fbExtDisableAF(
    Axis := axis3,
    Execute := bForceFall OR bEStopActive OR bNeedAxisReset
);

fbExtDisableYaw(
    Axis := axis4,
    Execute := bForceFall OR bEStopActive OR bNeedAxisReset
);

bExtBD := fbExtEnableBD.Enabled;
bExtAC := fbExtEnableAC.Enabled;
bExtAF := fbExtEnableAF.Enabled;
bExtYaw := fbExtEnableYaw.Enabled;

bRunForce := bForceMode
             AND bZeroDone
             AND bAxesReadyForForce
             AND axis1_power.Status
             AND Axis1_BrakeMotionOK
             AND axis2_power.Status
             AND axis3_power.Status
             AND axis4_power.Status
             AND bExtBD
             AND bExtAC
             AND bExtAF
             AND bExtYaw;

// 未进入实际力控运行（包括退出、急停、轴未就绪）时清除平面历史意图。
IF NOT bRunForce THEN
    bXIntent := FALSE;
    bZIntent := FALSE;
    bXDriveActive := FALSE;
    bZDriveActive := FALSE;
    Fx_work_target := 0.0;
    Fz_work_target := 0.0;
    Fx_work := 0.0;
    Fz_work := 0.0;
END_IF;


// =============================================================
// O. 编码器值 -> 机构学位置
// AC：-59 编码器对应 90°，编码器增大角度减小
// =============================================================
LBD_mm := BD_ActEnc + BD_KinOffset_mm;
LBD_m  := LBD_mm / 1000.0;

ThetaAC_deg := AC_ThetaRef_deg - (AC_ActEnc - AC_EncRef_deg);
ThetaAC_rad := ThetaAC_deg * DEG2RAD;


// =============================================================
// P. 当前 E 点正解
// =============================================================
bGeoOK := FALSE;

Cx := Ax0 + l_AC * COS(ThetaAC_rad);
Cz := Az0 + l_AC * SIN(ThetaAC_rad);

dxBC := Cx - Bx0;
dzBC := Cz - Bz0;
dBC := SQRT(dxBC * dxBC + dzBC * dzBC);

IF (LBD_m > 0.01) AND (dBC > 0.01) THEN
    IF (dBC < (LBD_m + l_CD - GeoMargin_m)) AND
       (dBC > (ABS(LBD_m - l_CD) + GeoMargin_m)) THEN

        alphaBC := F_Atan2_LREAL(y := dzBC, x := dxBC);
        cosBeta := (LBD_m * LBD_m + dBC * dBC - l_CD * l_CD) / (2.0 * LBD_m * dBC);

        IF (cosBeta <= 1.0) AND (cosBeta >= -1.0) THEN
            beta := ACOS(cosBeta);
            thBD := alphaBC - beta;

            Dx := Bx0 + LBD_m * COS(thBD);
            Dz := Bz0 + LBD_m * SIN(thBD);

            theta3 := F_Atan2_LREAL(y := Dz - Cz, x := Dx - Cx);

            // D 点不在 CE 上：D 相对 CE 垂直偏置 D_Offset_m
            // theta3 是 CD 方向，thetaCE 才是 CE 主杆方向
            IF l_CD > D_Offset_m THEN
                s_CD_CE := SQRT(l_CD * l_CD - D_Offset_m * D_Offset_m);
                gamma_DCE := ATAN(D_Offset_m / s_CD_CE);
                thetaCE := theta3 + CE_Sign * gamma_DCE;

                Ex := Cx + l_CE * COS(thetaCE);
                Ez := Cz + l_CE * SIN(thetaCE);

                bGeoOK := TRUE;
            END_IF;
        END_IF;
    END_IF;
END_IF;


// =============================================================
// Q. AC 机构角扰动 E 点正解
// =============================================================
bGeoOK_th := FALSE;

Cx_th := Ax0 + l_AC * COS(ThetaAC_rad + dTheta);
Cz_th := Az0 + l_AC * SIN(ThetaAC_rad + dTheta);

dxBC_th := Cx_th - Bx0;
dzBC_th := Cz_th - Bz0;
dBC_th := SQRT(dxBC_th * dxBC_th + dzBC_th * dzBC_th);

IF (LBD_m > 0.01) AND (dBC_th > 0.01) THEN
    IF (dBC_th < (LBD_m + l_CD - GeoMargin_m)) AND
       (dBC_th > (ABS(LBD_m - l_CD) + GeoMargin_m)) THEN

        alphaBC_th := F_Atan2_LREAL(y := dzBC_th, x := dxBC_th);
        cosBeta_th := (LBD_m * LBD_m + dBC_th * dBC_th - l_CD * l_CD) / (2.0 * LBD_m * dBC_th);

        IF (cosBeta_th <= 1.0) AND (cosBeta_th >= -1.0) THEN
            beta_th := ACOS(cosBeta_th);
            thBD_th := alphaBC_th - beta_th;

            Dx_th := Bx0 + LBD_m * COS(thBD_th);
            Dz_th := Bz0 + LBD_m * SIN(thBD_th);

            theta3_th := F_Atan2_LREAL(y := Dz_th - Cz_th, x := Dx_th - Cx_th);

            IF l_CD > D_Offset_m THEN
                s_CD_CE_th := SQRT(l_CD * l_CD - D_Offset_m * D_Offset_m);
                gamma_DCE_th := ATAN(D_Offset_m / s_CD_CE_th);
                thetaCE_th := theta3_th + CE_Sign * gamma_DCE_th;

                Ex_th := Cx_th + l_CE * COS(thetaCE_th);
                Ez_th := Cz_th + l_CE * SIN(thetaCE_th);

                bGeoOK_th := TRUE;
            END_IF;
        END_IF;
    END_IF;
END_IF;


// =============================================================
// R. BD 机构长度扰动 E 点正解
// =============================================================
bGeoOK_L := FALSE;

Cx_L := Cx;
Cz_L := Cz;

dxBC_L := Cx_L - Bx0;
dzBC_L := Cz_L - Bz0;
dBC_L := SQRT(dxBC_L * dxBC_L + dzBC_L * dzBC_L);

IF ((LBD_m + dL) > 0.01) AND (dBC_L > 0.01) THEN
    IF (dBC_L < ((LBD_m + dL) + l_CD - GeoMargin_m)) AND
       (dBC_L > (ABS((LBD_m + dL) - l_CD) + GeoMargin_m)) THEN

        alphaBC_L := F_Atan2_LREAL(y := dzBC_L, x := dxBC_L);
        cosBeta_L := ((LBD_m + dL) * (LBD_m + dL) + dBC_L * dBC_L - l_CD * l_CD)
                     / (2.0 * (LBD_m + dL) * dBC_L);

        IF (cosBeta_L <= 1.0) AND (cosBeta_L >= -1.0) THEN
            beta_L := ACOS(cosBeta_L);
            thBD_L := alphaBC_L - beta_L;

            Dx_L := Bx0 + (LBD_m + dL) * COS(thBD_L);
            Dz_L := Bz0 + (LBD_m + dL) * SIN(thBD_L);

            theta3_L := F_Atan2_LREAL(y := Dz_L - Cz_L, x := Dx_L - Cx_L);

            IF l_CD > D_Offset_m THEN
                s_CD_CE_L := SQRT(l_CD * l_CD - D_Offset_m * D_Offset_m);
                gamma_DCE_L := ATAN(D_Offset_m / s_CD_CE_L);
                thetaCE_L := theta3_L + CE_Sign * gamma_DCE_L;

                Ex_L := Cx_L + l_CE * COS(thetaCE_L);
                Ez_L := Cz_L + l_CE * SIN(thetaCE_L);

                bGeoOK_L := TRUE;
            END_IF;
        END_IF;
    END_IF;
END_IF;


// =============================================================
// S. E 点速度雅可比
// =============================================================
bValidJ := FALSE;
bSingular := FALSE;

IF bGeoOK AND bGeoOK_th AND bGeoOK_L THEN
    J11 := (Ex_th - Ex) / dTheta;
    J21 := (Ez_th - Ez) / dTheta;

    J12 := (Ex_L - Ex) / dL;
    J22 := (Ez_L - Ez) / dL;

    detJ := J11 * J22 - J12 * J21;

    IF ABS(detJ) > DetMin THEN
        bValidJ := TRUE;
    ELSE
        bSingular := TRUE;
    END_IF;
END_IF;


// =============================================================
// T. AC/BD 二维导纳 + 雅可比逆解
// 1) 平面 X/Z 导纳由显式欧拉改为一阶精确离散：M * dV/dt + B * V = F
//    Vss = Fadm / B
//    V(k+1) = Vss + (V(k)-Vss) * EXP(-B*Ts/M)
// 2) 撤力时使用 AdmB_Stop_X/Z 平滑衰减，轴减速度限幅约束最终命令。
// 3) VxyMax_mps = 0.300，先限制末端合速度，再做 J^-1。
// =============================================================
BD_Vraw_enc_s := 0.0;
AC_Vraw_enc_s := 0.0;
AF_Vraw_enc_s := 0.0;
Yaw_Vraw_enc_s := 0.0;

IF bRunForce AND bValidJ THEN
    Vx_last_mps := Vx_mps;
    Vz_last_mps := Vz_mps;

    // X 通道：有力用运动阻尼，撤力用停车阻尼。
    IF NOT bXDriveActive THEN
        AdmB_Use_X := AdmB_Stop_X;
        Fadm_X := 0.0;
    ELSE
        AdmB_Use_X := AdmB_Move_X;
        Fadm_X := ForceGain_X * TransWeight_X * Fx_work;
    END_IF;

    // Z 通道：有力用运动阻尼，撤力用停车阻尼。
    IF NOT bZDriveActive THEN
        AdmB_Use_Z := AdmB_Stop_Z;
        Fadm_Z := 0.0;
    ELSE
        AdmB_Use_Z := AdmB_Move_Z;
        Fadm_Z := ForceGain_Z * TransWeight_Z * Fz_work;
    END_IF;

    // M/B 安全保护，防止除零或负值。
    IF AdmM_X < 0.001 THEN
        AdmM_X_Use := 0.001;
    ELSE
        AdmM_X_Use := AdmM_X;
    END_IF;

    IF AdmM_Z < 0.001 THEN
        AdmM_Z_Use := 0.001;
    ELSE
        AdmM_Z_Use := AdmM_Z;
    END_IF;

    IF AdmB_Use_X < 0.001 THEN
        AdmB_X_UseSafe := 0.001;
    ELSE
        AdmB_X_UseSafe := AdmB_Use_X;
    END_IF;

    IF AdmB_Use_Z < 0.001 THEN
        AdmB_Z_UseSafe := 0.001;
    ELSE
        AdmB_Z_UseSafe := AdmB_Use_Z;
    END_IF;

    // 稳态速度。撤力时 Fadm=0，因此 Vss=0。
    Vxss_mps := Fadm_X / AdmB_X_UseSafe;
    Vzss_mps := Fadm_Z / AdmB_Z_UseSafe;

    // 精确离散指数项。
    IF Ts > 0.000001 THEN
        Vx_ExpK := EXP(-AdmB_X_UseSafe * Ts / AdmM_X_Use);
        Vz_ExpK := EXP(-AdmB_Z_UseSafe * Ts / AdmM_Z_Use);
    ELSE
        Vx_ExpK := 0.0;
        Vz_ExpK := 0.0;
    END_IF;

    Vx_mps := Vxss_mps + (Vx_last_mps - Vxss_mps) * Vx_ExpK;
    Vz_mps := Vzss_mps + (Vz_last_mps - Vzss_mps) * Vz_ExpK;

    IF Ts > 0.000001 THEN
        Ax_mps2 := (Vx_mps - Vx_last_mps) / Ts;
        Az_mps2 := (Vz_mps - Vz_last_mps) / Ts;
    ELSE
        Ax_mps2 := 0.0;
        Az_mps2 := 0.0;
    END_IF;

    // NaN / 极大值保护，避免后续 J^-1 或限幅触发 FPU invalid。
    IF Vx_mps <> Vx_mps THEN
        Vx_mps := 0.0;
        Vx_last_mps := 0.0;
        Ax_mps2 := 0.0;
    ELSIF ABS(Vx_mps) > Vplane_NumLimit_mps THEN
        Vx_mps := 0.0;
        Vx_last_mps := 0.0;
        Ax_mps2 := 0.0;
    END_IF;

    IF Vz_mps <> Vz_mps THEN
        Vz_mps := 0.0;
        Vz_last_mps := 0.0;
        Az_mps2 := 0.0;
    ELSIF ABS(Vz_mps) > Vplane_NumLimit_mps THEN
        Vz_mps := 0.0;
        Vz_last_mps := 0.0;
        Az_mps2 := 0.0;
    END_IF;

    // 限幅前理论平面速度。
    Vnorm_PreLimit_mps := SQRT(Vx_mps * Vx_mps + Vz_mps * Vz_mps);

    IF Vnorm_PreLimit_mps > VxyMax_mps THEN
        ScaleVel_Plane := VxyMax_mps / Vnorm_PreLimit_mps;
        Vx_mps := Vx_mps * ScaleVel_Plane;
        Vz_mps := Vz_mps * ScaleVel_Plane;
    ELSE
        ScaleVel_Plane := 1.0;
    END_IF;

    // 限幅后的真实平面速度。Watch 中 Vnorm 显示这个值。
    Vnorm_AfterLimit_mps := SQRT(Vx_mps * Vx_mps + Vz_mps * Vz_mps);
    Vnorm := Vnorm_AfterLimit_mps;

    qdotAC_rad_s := ( J22 * Vx_mps - J12 * Vz_mps) / detJ;
    qdotBD_m_s   := (-J21 * Vx_mps + J11 * Vz_mps) / detJ;

    // AC：机构角增大时，编码器减小。
    AC_Vraw_enc_s := -qdotAC_rad_s * RAD2DEG;

    // BD：1 mm = 1 mm，不做比例换算。
    BD_Vraw_enc_s := qdotBD_m_s * 1000.0;

ELSE
    Vx_mps := 0.0;
    Vz_mps := 0.0;
    Vx_last_mps := 0.0;
    Vz_last_mps := 0.0;

    Ax_mps2 := 0.0;
    Az_mps2 := 0.0;

    Vnorm_PreLimit_mps := 0.0;
    Vnorm_AfterLimit_mps := 0.0;
    Vnorm := 0.0;
    ScaleVel_Plane := 1.0;

    qdotAC_rad_s := 0.0;
    qdotBD_m_s := 0.0;
END_IF;

// axis3 AF 俯仰：Tz/Mz -> 俯仰角速度
// 本版关键修改：
// 1) 不再用显式欧拉 W += ((Madm-B*W)/J)*Ts 处理大 Stop 阻尼；
// 2) 改用一阶系统精确离散 W_new = Wss + (W_old-Wss)*EXP(-B*Ts/J)；
// 3) 撤力阻尼保持温和，减速由 AF_Dmax_enc_s2 最终约束。
IF bRunForce THEN
    AF_W_last_enc_s := AF_W_enc_s;

    bAF_TorqueActive := ABS(Mz_work_Nm) > 0.0001;

    IF bAF_TorqueActive THEN
        AdmB_Use_AF := AdmB_Move_AF;
        Madm_AF := TorqueGain_AF * Dir_Mz_AF * Mz_work_Nm;
    ELSE
        AdmB_Use_AF := AdmB_Stop_AF;
        Madm_AF := 0.0;
    END_IF;

    // 数值保护：J 和 B 都不允许过小。
    IF AdmJ_AF < 0.001 THEN
        AdmJ_AF_Use := 0.001;
    ELSE
        AdmJ_AF_Use := AdmJ_AF;
    END_IF;

    IF AdmB_Use_AF < 0.001 THEN
        AdmB_AF_UseSafe := 0.001;
    ELSE
        AdmB_AF_UseSafe := AdmB_Use_AF;
    END_IF;

    // 一阶导纳精确离散，撤力阻尼决定内部角速度衰减时间常数。
    IF Ts > 0.000001 THEN
        AF_ExpK := EXP(-AdmB_AF_UseSafe * Ts / AdmJ_AF_Use);
    ELSE
        AF_ExpK := 0.0;
    END_IF;

    AF_Wss_enc_s := Madm_AF / AdmB_AF_UseSafe;
    AF_W_enc_s := AF_Wss_enc_s + (AF_W_last_enc_s - AF_Wss_enc_s) * AF_ExpK;

    // 撤力后小速度直接归零，避免低速漂移。
    IF (NOT bAF_TorqueActive) AND (ABS(AF_W_enc_s) < AF_StopZeroVel_enc_s) THEN
        AF_W_enc_s := 0.0;
    END_IF;

    IF Ts > 0.000001 THEN
        AF_Alpha_enc_s2 := (AF_W_enc_s - AF_W_last_enc_s) / Ts;
    ELSE
        AF_Alpha_enc_s2 := 0.0;
    END_IF;

    // NaN / 极大值保护，避免再次触发 FPU invalid。
    IF AF_W_enc_s <> AF_W_enc_s THEN
        AF_W_enc_s := 0.0;
        AF_W_last_enc_s := 0.0;
        AF_Alpha_enc_s2 := 0.0;
    ELSIF ABS(AF_W_enc_s) > AF_NumLimit_enc_s THEN
        AF_W_enc_s := 0.0;
        AF_W_last_enc_s := 0.0;
        AF_Alpha_enc_s2 := 0.0;
    END_IF;

    AF_Vraw_enc_s := AF_W_enc_s;
ELSE
    AF_W_enc_s := 0.0;
    AF_W_last_enc_s := 0.0;
    AF_Alpha_enc_s2 := 0.0;
    AF_Vraw_enc_s := 0.0;
END_IF;

// axis4 底盘 yaw：稳定离散导纳
// 当前 yaw 主输入来自 FzYaw_work_N -> Myaw_work_Nm -> Mx_work_Nm。
// 这里继续使用 Mx_work_Nm 作为 yaw 有效输入，兼容你前面 Watch 变量。
IF bRunForce THEN
    Yaw_W_last_enc_s := Yaw_W_enc_s;

    YawInput_Nm := Mx_work_Nm;

    // 有 yaw 输入时用运动阻尼；撤力后用停车阻尼。
    IF ABS(YawInput_Nm) <= 0.0001 THEN
        AdmB_Use_Yaw := AdmB_Stop_Yaw;
        Madm_Yaw := 0.0;
    ELSE
        AdmB_Use_Yaw := AdmB_Move_Yaw;
        Madm_Yaw := TorqueGain_Yaw * Dir_Mx_Yaw * YawInput_Nm;
    END_IF;

    // J/B 安全保护。
    IF AdmJ_Yaw < 0.001 THEN
        AdmJ_Yaw_Use := 0.001;
    ELSE
        AdmJ_Yaw_Use := AdmJ_Yaw;
    END_IF;

    IF AdmB_Use_Yaw < 0.001 THEN
        AdmB_Yaw_UseSafe := 0.001;
    ELSE
        AdmB_Yaw_UseSafe := AdmB_Use_Yaw;
    END_IF;

    // 一阶导纳精确离散：
    // dW/dt = (Madm - B*W)/J
    // Wss = Madm/B
    // W(k+1) = Wss + (W(k)-Wss)*EXP(-B*Ts/J)
    Yaw_Wss_enc_s := Madm_Yaw / AdmB_Yaw_UseSafe;

    IF Ts > 0.000001 THEN
        Yaw_ExpK := EXP(-AdmB_Yaw_UseSafe * Ts / AdmJ_Yaw_Use);
    ELSE
        Yaw_ExpK := 0.0;
    END_IF;

    Yaw_W_enc_s :=
        Yaw_Wss_enc_s
      + (Yaw_W_last_enc_s - Yaw_Wss_enc_s) * Yaw_ExpK;

    IF Ts > 0.000001 THEN
        Yaw_Alpha_enc_s2 := (Yaw_W_enc_s - Yaw_W_last_enc_s) / Ts;
    ELSE
        Yaw_Alpha_enc_s2 := 0.0;
    END_IF;

    // NaN / 极大值保护，避免再次触发 FPU invalid。
    IF Yaw_W_enc_s <> Yaw_W_enc_s THEN
        Yaw_W_enc_s := 0.0;
        Yaw_W_last_enc_s := 0.0;
        Yaw_Alpha_enc_s2 := 0.0;
    ELSIF ABS(Yaw_W_enc_s) > Yaw_NumLimit_enc_s THEN
        Yaw_W_enc_s := 0.0;
        Yaw_W_last_enc_s := 0.0;
        Yaw_Alpha_enc_s2 := 0.0;
    END_IF;

    Yaw_Vraw_enc_s := Yaw_W_enc_s;
ELSE
    Yaw_W_enc_s := 0.0;
    Yaw_W_last_enc_s := 0.0;
    Yaw_Alpha_enc_s2 := 0.0;
    Yaw_Vraw_enc_s := 0.0;
END_IF;




// =============================================================
// T1. 机构学限位对力控 Vraw 的拦截
// 放在 U. 轴速度限幅之前；先判断，再进入速度/加速度/位置积分
// =============================================================
bLimitClampPlanar := FALSE;
bLimitClampAF := FALSE;

// BD 只受 CE-HI 限位
IF (BD_Vraw_enc_s > 0.0) AND bCEHI_Block_BD_Pos THEN
    BD_Vraw_enc_s := 0.0;
    bLimitClampPlanar := TRUE;
END_IF;

IF (BD_Vraw_enc_s < 0.0) AND bCEHI_Block_BD_Neg THEN
    BD_Vraw_enc_s := 0.0;
    bLimitClampPlanar := TRUE;
END_IF;

// AC 同时受 CAF 和 CE-HI 限位
IF (AC_Vraw_enc_s > 0.0) AND (bCAF_Block_AC_Pos OR bCEHI_Block_AC_Pos) THEN
    AC_Vraw_enc_s := 0.0;
    bLimitClampPlanar := TRUE;
END_IF;

IF (AC_Vraw_enc_s < 0.0) AND (bCAF_Block_AC_Neg OR bCEHI_Block_AC_Neg) THEN
    AC_Vraw_enc_s := 0.0;
    bLimitClampPlanar := TRUE;
END_IF;

// AF 同时受 CAF 和 CE-HI 限位
IF (AF_Vraw_enc_s > 0.0) AND (bCAF_Block_AF_Pos OR bCEHI_Block_AF_Pos) THEN
    AF_Vraw_enc_s := 0.0;
    bLimitClampAF := TRUE;
END_IF;

IF (AF_Vraw_enc_s < 0.0) AND (bCAF_Block_AF_Neg OR bCEHI_Block_AF_Neg) THEN
    AF_Vraw_enc_s := 0.0;
    bLimitClampAF := TRUE;
END_IF;

// 清导纳内部速度记忆，防止继续顶限位
IF bLimitClampPlanar THEN
    Vx_mps := 0.0;
    Vz_mps := 0.0;
    Vx_last_mps := 0.0;
    Vz_last_mps := 0.0;
    Ax_mps2 := 0.0;
    Az_mps2 := 0.0;
END_IF;

IF bLimitClampAF THEN
    AF_W_enc_s := 0.0;
    AF_W_last_enc_s := 0.0;
    AF_Alpha_enc_s2 := 0.0;
END_IF;


// =============================================================
// U. 轴速度限幅
// =============================================================
ScaleVel := 1.0;
ScaleVel_Axis := 1.0;

IF ABS(BD_Vraw_enc_s) > BD_Vmax_enc_s THEN
    tmpScale := BD_Vmax_enc_s / ABS(BD_Vraw_enc_s);
    IF tmpScale < ScaleVel THEN
        ScaleVel := tmpScale;
    END_IF;
END_IF;

IF ABS(AC_Vraw_enc_s) > AC_Vmax_enc_s THEN
    tmpScale := AC_Vmax_enc_s / ABS(AC_Vraw_enc_s);
    IF tmpScale < ScaleVel THEN
        ScaleVel := tmpScale;
    END_IF;
END_IF;

ScaleVel_Axis := ScaleVel;

BD_Vraw_enc_s := BD_Vraw_enc_s * ScaleVel_Axis;
AC_Vraw_enc_s := AC_Vraw_enc_s * ScaleVel_Axis;

// AF/Yaw 速度限幅：不用 x/ABS(x)，避免 Infinity/Infinity 触发 FPU invalid。
IF AF_Vraw_enc_s <> AF_Vraw_enc_s THEN
    AF_Vraw_enc_s := 0.0;
    AF_W_enc_s := 0.0;
    AF_W_last_enc_s := 0.0;
ELSIF ABS(AF_Vraw_enc_s) > AF_NumLimit_enc_s THEN
    AF_Vraw_enc_s := 0.0;
    AF_W_enc_s := 0.0;
    AF_W_last_enc_s := 0.0;
END_IF;

IF AF_Vraw_enc_s > AF_Vmax_enc_s THEN
    AF_Vraw_enc_s := AF_Vmax_enc_s;
ELSIF AF_Vraw_enc_s < -AF_Vmax_enc_s THEN
    AF_Vraw_enc_s := -AF_Vmax_enc_s;
END_IF;

IF Yaw_Vraw_enc_s <> Yaw_Vraw_enc_s THEN
    Yaw_Vraw_enc_s := 0.0;
    Yaw_W_enc_s := 0.0;
    Yaw_W_last_enc_s := 0.0;
ELSIF ABS(Yaw_Vraw_enc_s) > 100000.0 THEN
    Yaw_Vraw_enc_s := 0.0;
    Yaw_W_enc_s := 0.0;
    Yaw_W_last_enc_s := 0.0;
END_IF;

IF Yaw_Vraw_enc_s > Yaw_Vmax_enc_s THEN
    Yaw_Vraw_enc_s := Yaw_Vmax_enc_s;
ELSIF Yaw_Vraw_enc_s < -Yaw_Vmax_enc_s THEN
    Yaw_Vraw_enc_s := -Yaw_Vmax_enc_s;
END_IF;


// =============================================================
// V. 加速度限幅
// =============================================================
BD_Vlast_enc_s := BD_Vcmd_enc_s;
AC_Vlast_enc_s := AC_Vcmd_enc_s;
AF_Vlast_enc_s := AF_Vcmd_enc_s;
Yaw_Vlast_enc_s := Yaw_Vcmd_enc_s;

// AC/BD 加减速度限幅：
// 1) 加速使用 BD_Amax/AC_Amax；
// 2) 撤力减速或反向使用 BD_Dmax/AC_Dmax；
// 3) 最后用同一个 ScaleAcc_Axis 同步缩放 BD/AC，保持末端方向不被破坏。
BD_dV_enc_s := BD_Vraw_enc_s - BD_Vlast_enc_s;
AC_dV_enc_s := AC_Vraw_enc_s - AC_Vlast_enc_s;

IF (ABS(BD_Vraw_enc_s) < ABS(BD_Vlast_enc_s)) OR (BD_Vraw_enc_s * BD_Vlast_enc_s < 0.0) THEN
    BD_dVmax_enc_s := BD_Dmax_enc_s2 * Ts;
ELSE
    BD_dVmax_enc_s := BD_Amax_enc_s2 * Ts;
END_IF;

IF (ABS(AC_Vraw_enc_s) < ABS(AC_Vlast_enc_s)) OR (AC_Vraw_enc_s * AC_Vlast_enc_s < 0.0) THEN
    AC_dVmax_enc_s := AC_Dmax_enc_s2 * Ts;
ELSE
    AC_dVmax_enc_s := AC_Amax_enc_s2 * Ts;
END_IF;

ScaleAcc := 1.0;
ScaleAcc_Axis := 1.0;

IF ABS(BD_dV_enc_s) > BD_dVmax_enc_s THEN
    IF BD_dVmax_enc_s > 0.0 THEN
        tmpScale := BD_dVmax_enc_s / ABS(BD_dV_enc_s);
    ELSE
        tmpScale := 0.0;
    END_IF;
    IF tmpScale < ScaleAcc THEN
        ScaleAcc := tmpScale;
    END_IF;
END_IF;

IF ABS(AC_dV_enc_s) > AC_dVmax_enc_s THEN
    IF AC_dVmax_enc_s > 0.0 THEN
        tmpScale := AC_dVmax_enc_s / ABS(AC_dV_enc_s);
    ELSE
        tmpScale := 0.0;
    END_IF;
    IF tmpScale < ScaleAcc THEN
        ScaleAcc := tmpScale;
    END_IF;
END_IF;

ScaleAcc_Axis := ScaleAcc;

BD_Vcmd_enc_s := BD_Vlast_enc_s + BD_dV_enc_s * ScaleAcc_Axis;
AC_Vcmd_enc_s := AC_Vlast_enc_s + AC_dV_enc_s * ScaleAcc_Axis;

IF Ts > 0.000001 THEN
    BD_Acmd_enc_s2 := (BD_Vcmd_enc_s - BD_Vlast_enc_s) / Ts;
    AC_Acmd_enc_s2 := (AC_Vcmd_enc_s - AC_Vlast_enc_s) / Ts;
ELSE
    BD_Acmd_enc_s2 := 0.0;
    AC_Acmd_enc_s2 := 0.0;
END_IF;

// AF 加减速度限幅：加速用 AF_Amax，撤力减速/反向用更大的 AF_Dmax。
AF_dV_enc_s := AF_Vraw_enc_s - AF_Vlast_enc_s;

IF (ABS(AF_Vraw_enc_s) < ABS(AF_Vlast_enc_s)) OR (AF_Vraw_enc_s * AF_Vlast_enc_s < 0.0) THEN
    AF_dVmax_enc_s := AF_Dmax_enc_s2 * Ts;
ELSE
    AF_dVmax_enc_s := AF_Amax_enc_s2 * Ts;
END_IF;

IF AF_dV_enc_s > AF_dVmax_enc_s THEN
    AF_dV_enc_s := AF_dVmax_enc_s;
ELSIF AF_dV_enc_s < -AF_dVmax_enc_s THEN
    AF_dV_enc_s := -AF_dVmax_enc_s;
END_IF;

AF_Vcmd_enc_s := AF_Vlast_enc_s + AF_dV_enc_s;

IF Ts > 0.000001 THEN
    AF_Acmd_enc_s2 := (AF_Vcmd_enc_s - AF_Vlast_enc_s) / Ts;
ELSE
    AF_Acmd_enc_s2 := 0.0;
END_IF;

// yaw 加减速度限幅：加速用 Yaw_Amax，撤力减速/反向用 Yaw_Dmax。
Yaw_dV_enc_s := Yaw_Vraw_enc_s - Yaw_Vlast_enc_s;

IF (ABS(Yaw_Vraw_enc_s) < ABS(Yaw_Vlast_enc_s)) OR (Yaw_Vraw_enc_s * Yaw_Vlast_enc_s < 0.0) THEN
    Yaw_dVmax_enc_s := Yaw_Dmax_enc_s2 * Ts;
ELSE
    Yaw_dVmax_enc_s := Yaw_Amax_enc_s2 * Ts;
END_IF;

IF Yaw_dV_enc_s > Yaw_dVmax_enc_s THEN
    Yaw_dV_enc_s := Yaw_dVmax_enc_s;
ELSIF Yaw_dV_enc_s < -Yaw_dVmax_enc_s THEN
    Yaw_dV_enc_s := -Yaw_dVmax_enc_s;
END_IF;

Yaw_Vcmd_enc_s := Yaw_Vlast_enc_s + Yaw_dV_enc_s;

IF Ts > 0.000001 THEN
    Yaw_Acmd_enc_s2 := (Yaw_Vcmd_enc_s - Yaw_Vlast_enc_s) / Ts;
ELSE
    Yaw_Acmd_enc_s2 := 0.0;
END_IF;




// =============================================================
// V1. 机构学限位对力控 Vcmd 的最终保险
// 放在 W. 小速度归零之前，位置积分之前
// =============================================================
// BD
IF (BD_Vcmd_enc_s > 0.0) AND bCEHI_Block_BD_Pos THEN
    BD_Vcmd_enc_s := 0.0;
    BD_Acmd_enc_s2 := 0.0;
END_IF;

IF (BD_Vcmd_enc_s < 0.0) AND bCEHI_Block_BD_Neg THEN
    BD_Vcmd_enc_s := 0.0;
    BD_Acmd_enc_s2 := 0.0;
END_IF;

// AC
IF (AC_Vcmd_enc_s > 0.0) AND (bCAF_Block_AC_Pos OR bCEHI_Block_AC_Pos) THEN
    AC_Vcmd_enc_s := 0.0;
    AC_Acmd_enc_s2 := 0.0;
END_IF;

IF (AC_Vcmd_enc_s < 0.0) AND (bCAF_Block_AC_Neg OR bCEHI_Block_AC_Neg) THEN
    AC_Vcmd_enc_s := 0.0;
    AC_Acmd_enc_s2 := 0.0;
END_IF;

// AF
IF (AF_Vcmd_enc_s > 0.0) AND (bCAF_Block_AF_Pos OR bCEHI_Block_AF_Pos) THEN
    AF_Vcmd_enc_s := 0.0;
    AF_Acmd_enc_s2 := 0.0;
    AF_W_enc_s := 0.0;
    AF_W_last_enc_s := 0.0;
END_IF;

IF (AF_Vcmd_enc_s < 0.0) AND (bCAF_Block_AF_Neg OR bCEHI_Block_AF_Neg) THEN
    AF_Vcmd_enc_s := 0.0;
    AF_Acmd_enc_s2 := 0.0;
    AF_W_enc_s := 0.0;
    AF_W_last_enc_s := 0.0;
END_IF;


// =============================================================
// W. 小速度归零
// =============================================================
IF ABS(BD_Vcmd_enc_s) < 0.001 THEN
    BD_Vcmd_enc_s := 0.0;
END_IF;

IF ABS(AC_Vcmd_enc_s) < 0.001 THEN
    AC_Vcmd_enc_s := 0.0;
END_IF;

IF ABS(AF_Vcmd_enc_s) < 0.02 THEN
    AF_Vcmd_enc_s := 0.0;
END_IF;

IF ABS(Yaw_Vcmd_enc_s) < 0.001 THEN
    Yaw_Vcmd_enc_s := 0.0;
END_IF;

// =============================================================
// W1. 轴1抱闸未释放时冻结 BD 给定
// 防止抱闸合上或释放延时未到时，BD 外部位置继续积分。
// =============================================================
IF NOT Axis1_BrakeMotionOK THEN
    BD_Vraw_enc_s := 0.0;
    BD_Vcmd_enc_s := 0.0;
    BD_Vlast_enc_s := 0.0;
    BD_Acmd_enc_s2 := 0.0;
    qdotBD_m_s := 0.0;
    BD_PosCmd_Enc := BD_ActEnc;
END_IF;


// =============================================================
// X. 力控基础软限位
// 当前只对 axis1=BD 编码器 2~600 做限位
// =============================================================
bForceSoftLimit := FALSE;

BD_NextCmd_Enc := BD_PosCmd_Enc + BD_Vcmd_enc_s * Ts;
AC_NextCmd_Enc := AC_PosCmd_Enc + AC_Vcmd_enc_s * Ts;
AF_NextCmd_Enc := AF_PosCmd_Enc + AF_Vcmd_enc_s * Ts;
Yaw_NextCmd_Enc := Yaw_PosCmd_Enc + Yaw_Vcmd_enc_s * Ts;

IF (BD_NextCmd_Enc < BD_EncMin) OR (BD_NextCmd_Enc > BD_EncMax) THEN
    bForceSoftLimit := TRUE;
END_IF;

IF bUseAFLimit THEN
    IF (AF_NextCmd_Enc < AF_EncMin) OR (AF_NextCmd_Enc > AF_EncMax) THEN
        bForceSoftLimit := TRUE;
    END_IF;
END_IF;

IF (Yaw_NextCmd_Enc < Base_EncMin) OR (Yaw_NextCmd_Enc > Base_EncMax) THEN
    bForceSoftLimit := TRUE;
END_IF;

IF bForceSoftLimit THEN
    BD_Vcmd_enc_s := 0.0;
    AC_Vcmd_enc_s := 0.0;
    AF_Vcmd_enc_s := 0.0;
    Yaw_Vcmd_enc_s := 0.0;

    BD_Acmd_enc_s2 := 0.0;
    AC_Acmd_enc_s2 := 0.0;
    AF_Acmd_enc_s2 := 0.0;
    Yaw_Acmd_enc_s2 := 0.0;

    Vx_mps := 0.0;
    Vz_mps := 0.0;
    AF_W_enc_s := 0.0;
    Yaw_W_enc_s := 0.0;
END_IF;


// =============================================================
// Y. 位置积分
// 外部位置给定使用真实 NC 编码器坐标
// =============================================================
IF bRunForce AND NOT bForceSoftLimit THEN
    BD_PosCmd_Enc := BD_PosCmd_Enc + BD_Vcmd_enc_s * Ts;
    AC_PosCmd_Enc := AC_PosCmd_Enc + AC_Vcmd_enc_s * Ts;
    AF_PosCmd_Enc := AF_PosCmd_Enc + AF_Vcmd_enc_s * Ts;
    Yaw_PosCmd_Enc := Yaw_PosCmd_Enc + Yaw_Vcmd_enc_s * Ts;
END_IF;


// =============================================================
// Z. Direction 判断
// =============================================================
IF BD_Vcmd_enc_s > 0.001 THEN
    DirBD := 1;
ELSIF BD_Vcmd_enc_s < -0.001 THEN
    DirBD := -1;
ELSE
    DirBD := 0;
END_IF;

IF AC_Vcmd_enc_s > 0.001 THEN
    DirAC := 1;
ELSIF AC_Vcmd_enc_s < -0.001 THEN
    DirAC := -1;
ELSE
    DirAC := 0;
END_IF;

IF AF_Vcmd_enc_s > 0.001 THEN
    DirAF := 1;
ELSIF AF_Vcmd_enc_s < -0.001 THEN
    DirAF := -1;
ELSE
    DirAF := 0;
END_IF;

IF Yaw_Vcmd_enc_s > 0.001 THEN
    DirYaw := 1;
ELSIF Yaw_Vcmd_enc_s < -0.001 THEN
    DirYaw := -1;
ELSE
    DirYaw := 0;
END_IF;


// =============================================================
// Z1. 每周期 Feed axis1 / axis2 / axis3 / axis4
// 急停、未 Ready、未力控时，不再 Feed，避免恢复后继续追旧目标。
// =============================================================
IF bRunForce AND bAxesReadyForForce THEN
    bFeedBD := MC_ExtSetPointGenFeed(
        Axis := axis1,
        Position := BD_PosCmd_Enc,
        Velocity := ABS(BD_Vcmd_enc_s),
        Acceleration := ABS(BD_Acmd_enc_s2),
        Direction := DirBD
    );

    bFeedAC := MC_ExtSetPointGenFeed(
        Axis := axis2,
        Position := AC_PosCmd_Enc,
        Velocity := ABS(AC_Vcmd_enc_s),
        Acceleration := ABS(AC_Acmd_enc_s2),
        Direction := DirAC
    );

    bFeedAF := MC_ExtSetPointGenFeed(
        Axis := axis3,
        Position := AF_PosCmd_Enc,
        Velocity := ABS(AF_Vcmd_enc_s),
        Acceleration := ABS(AF_Acmd_enc_s2),
        Direction := DirAF
    );

    bFeedYaw := MC_ExtSetPointGenFeed(
        Axis := axis4,
        Position := Yaw_PosCmd_Enc,
        Velocity := ABS(Yaw_Vcmd_enc_s),
        Acceleration := ABS(Yaw_Acmd_enc_s2),
        Direction := DirYaw
    );
ELSE
    bFeedBD := FALSE;
    bFeedAC := FALSE;
    bFeedAF := FALSE;
    bFeedYaw := FALSE;

    // 非力控/急停/轴未 Ready 时保持目标等于当前位置，防止恢复后跳变。
    IF NOT bRunForce THEN
        BD_PosCmd_Enc := BD_ActEnc;
        AC_PosCmd_Enc := AC_ActEnc;
        AF_PosCmd_Enc := AF_ActEnc;
        Yaw_PosCmd_Enc := Yaw_ActEnc;
    END_IF;
END_IF;


// =============================================================
// Z2. 抱闸和灯
// =============================================================
// 轴1抱闸 axis1baozha 已在 D1 中按“轴1真实使能 + 无故障 + 300ms 延时”逻辑处理。
// 这里保留 axis4 原逻辑。注意：axis4 不受 CE-HI 限位影响。
axis4baozha := ballow_axis4jogfw OR ballow_axis4jogbw OR bRunForce;

// 电磁阀和电磁阀灯完全独立，不经过 CAF/CEHI 限位。
valveopen1 := valvejudge;
valveopen2 := valvejudge;
valvelight := valvejudge;

// 指示灯也从 CEHI/CAF 限位逻辑中拆出来：
// 手动模式下，只要按钮输入为 TRUE 就亮，用于确认按钮链路；
// 力控模式下，对应轴有速度给定时也亮。
// 这样即使某方向被软限位禁止，按键灯仍能亮，便于判断“输入有效但被限位拦截”。
bOutput_axis1light :=
    bInput_axis1jogfw OR bInput_axis1jogbw
    OR (bRunForce AND (ABS(BD_Vcmd_enc_s) > 0.001));

bOutput_axis2light :=
    bInput_axis2jogfw OR bInput_axis2jogbw
    OR (bRunForce AND (ABS(AC_Vcmd_enc_s) > 0.001));

bOutput_axis3light :=
    bInput_axis3jogfw OR bInput_axis3jogbw
    OR (bRunForce AND (ABS(AF_Vcmd_enc_s) > 0.02));

bOutput_axis4light :=
    bInput_axis4jogfw OR bInput_axis4jogbw
    OR (bRunForce AND (ABS(Yaw_Vcmd_enc_s) > 0.001));

    likonglight := bForceMode;

// =============================================================
// Z3. 错误输出
// =============================================================
axis1_status(Axis := axis1, Enable := TRUE);
axis2_status(Axis := axis2, Enable := TRUE);
axis3_status(Axis := axis3, Enable := TRUE);
axis4_status(Axis := axis4, Enable := TRUE);

bAxis1Err := axis1_power.Error OR axis1_status.Error OR axis1_status.ErrorStop;
bAxis2Err := axis2_power.Error OR axis2_status.Error OR axis2_status.ErrorStop;
bAxis3Err := axis3_power.Error OR axis3_status.Error OR axis3_status.ErrorStop;
bAxis4Err := axis4_power.Error OR axis4_status.Error OR axis4_status.ErrorStop;

bAnyAxisErr := bAxis1Err OR bAxis2Err OR bAxis3Err OR bAxis4Err;

IF bResetStopReason THEN
    StopReasonCode := 0;
    bStopReasonLatched := FALSE;
END_IF;

IF bRunForce AND NOT bStopReasonLatched THEN

    IF NOT bForceMode THEN
        StopReasonCode := 1;
        bStopReasonLatched := TRUE;

    ELSIF NOT bAxesReadyForForce THEN
        StopReasonCode := 2;
        bStopReasonLatched := TRUE;

   ELSIF bAnyAxisErr THEN
    StopReasonCode := 3;
    bStopReasonLatched := TRUE;
    

    ELSIF bCEHI_Block_BD_Pos OR bCEHI_Block_BD_Neg
       OR bCEHI_Block_AC_Pos OR bCEHI_Block_AC_Neg
       OR bCEHI_Block_AF_Pos OR bCEHI_Block_AF_Neg THEN
        StopReasonCode := 4;
        bStopReasonLatched := TRUE;

    ELSIF bCAF_Block_AC_Pos OR bCAF_Block_AC_Neg
       OR bCAF_Block_AF_Pos OR bCAF_Block_AF_Neg THEN
        StopReasonCode := 5;
        bStopReasonLatched := TRUE;

    ELSIF NOT bExtBD OR NOT bExtAC THEN
        StopReasonCode := 6;
        bStopReasonLatched := TRUE;

    ELSIF NOT Axis1_BrakeMotionOK THEN
        StopReasonCode := 7;
        bStopReasonLatched := TRUE;
    END_IF;

END_IF;

bError := axis1_power.Error OR axis2_power.Error OR axis3_power.Error OR axis4_power.Error
       OR axis1_jogerror OR axis2_jogerror OR axis3_jogerror OR axis4_jogerror
       OR fbExtEnableBD.Error OR fbExtEnableAC.Error OR fbExtEnableAF.Error OR fbExtEnableYaw.Error
       OR fbExtDisableBD.Error OR fbExtDisableAC.Error OR fbExtDisableAF.Error OR fbExtDisableYaw.Error
       OR axis1_reset.Error OR axis2_reset.Error OR axis3_reset.Error OR axis4_reset.Error;

IF axis1_power.Error THEN
    nErrorID := axis1_power.ErrorID;
ELSIF axis2_power.Error THEN
    nErrorID := axis2_power.ErrorID;
ELSIF axis3_power.Error THEN
    nErrorID := axis3_power.ErrorID;
ELSIF axis4_power.Error THEN
    nErrorID := axis4_power.ErrorID;
ELSIF axis1_jogerror THEN
    nErrorID := axis1_jogerrorid;
ELSIF axis2_jogerror THEN
    nErrorID := axis2_jogerrorid;
ELSIF axis3_jogerror THEN
    nErrorID := axis3_jogerrorid;
ELSIF axis4_jogerror THEN
    nErrorID := axis4_jogerrorid;
ELSIF fbExtEnableBD.Error THEN
    nErrorID := fbExtEnableBD.ErrorID;
ELSIF fbExtEnableAC.Error THEN
    nErrorID := fbExtEnableAC.ErrorID;
ELSIF fbExtEnableAF.Error THEN
    nErrorID := fbExtEnableAF.ErrorID;
ELSIF fbExtEnableYaw.Error THEN
    nErrorID := fbExtEnableYaw.ErrorID;
ELSIF fbExtDisableBD.Error THEN
    nErrorID := fbExtDisableBD.ErrorID;
ELSIF fbExtDisableAC.Error THEN
    nErrorID := fbExtDisableAC.ErrorID;
ELSIF fbExtDisableAF.Error THEN
    nErrorID := fbExtDisableAF.ErrorID;
ELSIF fbExtDisableYaw.Error THEN
    nErrorID := fbExtDisableYaw.ErrorID;
ELSIF axis1_reset.Error THEN
    nErrorID := axis1_reset.ErrorID;
ELSIF axis2_reset.Error THEN
    nErrorID := axis2_reset.ErrorID;
ELSIF axis3_reset.Error THEN
    nErrorID := axis3_reset.ErrorID;
ELSIF axis4_reset.Error THEN
    nErrorID := axis4_reset.ErrorID;
ELSE
    nErrorID := 0;
END_IF;

END_PROGRAM

// ---- POUs/FB_Calc_CEHI_Geo.TcPOU

// =============================================================
// FUNCTION_BLOCK：FB_Calc_CEHI_Geo
// MATLAB 对应关系：
//   res.F = A + l_AF*[cos(th_af); sin(th_af)]
//   res.G = C + (res.F - A)
//   th_CH = th_af - angle_GCH
//   res.H = C + l_CH*[cos(th_CH); sin(th_CH)]
//   res.I = E + (res.H - res.C)
// 这里不显式输出 F/G，但按照同一逻辑构造 thetaAF_abs 与 thetaCH/EI。
// =============================================================
FUNCTION_BLOCK FB_Calc_CEHI_Geo
VAR_INPUT
    BD_Enc_mm             : LREAL;
    AC_Enc_deg            : LREAL;
    AF_Enc_deg            : LREAL;

    BD_KinOffset_mm       : LREAL;

    AC_EncRef_deg         : LREAL;
    AC_ThetaRef_deg       : LREAL;

    Ax0                   : LREAL;
    Az0                   : LREAL;
    Bx0                   : LREAL;
    Bz0                   : LREAL;

    l_AC_m                : LREAL;
    l_CD_m                : LREAL;
    l_CE_m                : LREAL;
    qOffset_m             : LREAL;
    l_CH_m                : LREAL;

    BD_BRANCH             : LREAL;     // -1：thetaBD = alphaBC - beta；+1：thetaBD = alphaBC + beta
    CE_SIGN               : LREAL;     // +1 / -1，D/q 偏置到 CE 方向的装配符号

    AF_HorizontalEnc_deg  : LREAL;
    AF_CHOffset_deg       : LREAL;     // AF=水平时 EI/CH 与 +X 的夹角，当前保持 MAIN 中最新值 15 deg
    AF_EncDir_CH          : LREAL;     // 当前保持 MAIN 中最新值 -1：thetaEI = 205 - AF + offset

    GeoMargin_m           : LREAL;
END_VAR
VAR_OUTPUT
    Valid                 : BOOL;
    ErrorID               : INT;

    Cx                    : LREAL;
    Cz                    : LREAL;
    Dx                    : LREAL;
    Dz                    : LREAL;
    Qx                    : LREAL;
    Qz                    : LREAL;
    Ex                    : LREAL;
    Ez                    : LREAL;

    Hx                    : LREAL;
    Hz                    : LREAL;
    Ix                    : LREAL;
    Iz                    : LREAL;

    thetaCE_rad           : LREAL;
    ThetaCH_rad           : LREAL;
    ThetaCH_deg           : LREAL;
    ThetaAF_abs_deg       : LREAL;     // 新增诊断：按 MATLAB th_af 含义得到的 AF 绝对角
    DeltaCH_CE_deg        : LREAL;

    uCEx                  : LREAL;
    uCEz                  : LREAL;

    CEHI_Dis_m            : LREAL;
    CEHI_DisSigned_m      : LREAL;
    DisFromH_m            : LREAL;
    DisFromI_m            : LREAL;
    DisFromHIAvg_m        : LREAL;
    DisDiff_m             : LREAL;

    CE_L_Check_m          : LREAL;
    Q_Offset_Check_m      : LREAL;
    CH_L_Check_m          : LREAL;
    EI_L_Check_m          : LREAL;
    HI_L_Check_m          : LREAL;
    HI_ParallelErr_m      : LREAL;
END_VAR
VAR
    LBD_m        : LREAL;

    ThetaAC_deg  : LREAL;
    ThetaAC_rad  : LREAL;

    dxBC         : LREAL;
    dzBC         : LREAL;
    dBC          : LREAL;

    alphaBC      : LREAL;
    cosBeta      : LREAL;
    beta         : LREAL;
    thBD         : LREAL;

    thetaCD      : LREAL;
    s_CD_CE      : LREAL;
    gamma_DCE    : LREAL;

    uCHx         : LREAL;
    uCHz         : LREAL;

    // MATLAB 中 th_af - angle_GCH。这里 angle_GCH 取 90 度三角板关系，
    // 因此 thetaCH = thetaAF_abs - 90 = thetaEI。
    GCH_Matlab_deg : LREAL := 90.0;

    DEG2RAD_local : LREAL := 0.0174532925199433;
    RAD2DEG_local : LREAL := 57.29577951308232;
END_VAR



// 默认无效
Valid := FALSE;
ErrorID := 0;

Cx := 0.0; Cz := 0.0;
Dx := 0.0; Dz := 0.0;
Qx := 0.0; Qz := 0.0;
Ex := 0.0; Ez := 0.0;
Hx := 0.0; Hz := 0.0;
Ix := 0.0; Iz := 0.0;

thetaCE_rad := 0.0;
ThetaCH_rad := 0.0;
ThetaCH_deg := 0.0;
ThetaAF_abs_deg := 0.0;
DeltaCH_CE_deg := 0.0;

uCEx := 1.0;
uCEz := 0.0;

CEHI_Dis_m := -1.0;
CEHI_DisSigned_m := 0.0;
DisFromH_m := -1.0;
DisFromI_m := -1.0;
DisFromHIAvg_m := -1.0;
DisDiff_m := 0.0;

CE_L_Check_m := 0.0;
Q_Offset_Check_m := 0.0;
CH_L_Check_m := 0.0;
EI_L_Check_m := 0.0;
HI_L_Check_m := 0.0;
HI_ParallelErr_m := 0.0;

// BD 编码器 -> 机构长度
LBD_m := (BD_Enc_mm + BD_KinOffset_mm) / 1000.0;

// AC 编码器 -> AC 机构角
ThetaAC_deg := AC_ThetaRef_deg - (AC_Enc_deg - AC_EncRef_deg);
ThetaAC_rad := ThetaAC_deg * DEG2RAD_local;

// C 点
Cx := Ax0 + l_AC_m * COS(ThetaAC_rad);
Cz := Az0 + l_AC_m * SIN(ThetaAC_rad);

// B-C
dxBC := Cx - Bx0;
dzBC := Cz - Bz0;
dBC  := SQRT(dxBC * dxBC + dzBC * dzBC);

IF (LBD_m <= 0.01) OR (dBC <= 0.01) THEN
    ErrorID := 1;
    RETURN;
END_IF;

IF NOT ((dBC < (LBD_m + l_CD_m - GeoMargin_m)) AND
        (dBC > (ABS(LBD_m - l_CD_m) + GeoMargin_m))) THEN
    ErrorID := 2;
    RETURN;
END_IF;

// 三角形 B-C-D。这里保留 PLC 的 BD_BRANCH，用你的最新参数 -1。
alphaBC := F_Atan2_LREAL(y := dzBC, x := dxBC);

cosBeta := (LBD_m * LBD_m + dBC * dBC - l_CD_m * l_CD_m)
           / (2.0 * LBD_m * dBC);

IF cosBeta > 1.0 THEN
    cosBeta := 1.0;
ELSIF cosBeta < -1.0 THEN
    cosBeta := -1.0;
END_IF;

beta := ACOS(cosBeta);
thBD := alphaBC + BD_BRANCH * beta;

Dx := Bx0 + LBD_m * COS(thBD);
Dz := Bz0 + LBD_m * SIN(thBD);

// CD 方向
thetaCD := F_Atan2_LREAL(y := Dz - Cz, x := Dx - Cx);

// D 到 CE 的垂直偏置 qOffset_m。MATLAB 原代码没有这一步，PLC 保留。
IF l_CD_m <= ABS(qOffset_m) THEN
    ErrorID := 3;
    RETURN;
END_IF;

s_CD_CE := SQRT(l_CD_m * l_CD_m - qOffset_m * qOffset_m);
gamma_DCE := ATAN(qOffset_m / s_CD_CE);

thetaCE_rad := thetaCD + CE_SIGN * gamma_DCE;

uCEx := COS(thetaCE_rad);
uCEz := SIN(thetaCE_rad);

// Q 点：D 到 CE 的垂足
Qx := Cx + s_CD_CE * uCEx;
Qz := Cz + s_CD_CE * uCEz;

// CE 末端 E
Ex := Cx + l_CE_m * uCEx;
Ez := Cz + l_CE_m * uCEz;

// =============================================================
// 后级 H/I：按 MATLAB 机构方法写清楚
// AF=水平时，EI/CH 与 +X 的夹角为 AF_CHOffset_deg。
// AF 减小时，若 AF_EncDir_CH=-1，则 EI/CH 角度增大。
// thetaAF_abs 只是诊断量；真正用于 H/I 的是 thetaCH = thetaAF_abs - 90。
// =============================================================
ThetaCH_deg := AF_EncDir_CH * (AF_Enc_deg - AF_HorizontalEnc_deg) + AF_CHOffset_deg;
ThetaAF_abs_deg := ThetaCH_deg + GCH_Matlab_deg;
ThetaCH_deg := ThetaAF_abs_deg - GCH_Matlab_deg;
ThetaCH_rad := ThetaCH_deg * DEG2RAD_local;

uCHx := COS(ThetaCH_rad);
uCHz := SIN(ThetaCH_rad);

// MATLAB：H = C + l_CH*[cos(th_CH), sin(th_CH)]
Hx := Cx + l_CH_m * uCHx;
Hz := Cz + l_CH_m * uCHz;

// MATLAB：I = E + (H - C)，从而 HI 与 CE 平行
Ix := Ex + (Hx - Cx);
Iz := Ez + (Hz - Cz);

// H/I 到 CE 直线的有符号距离。CE 直线以 C 为基点，方向 uCE。
CEHI_DisSigned_m := uCEx * (Hz - Cz) - uCEz * (Hx - Cx);

DisFromH_m := ABS(
    uCEx * (Hz - Cz) - uCEz * (Hx - Cx)
);

DisFromI_m := ABS(
    uCEx * (Iz - Cz) - uCEz * (Ix - Cx)
);

DisFromHIAvg_m := 0.5 * (DisFromH_m + DisFromI_m);
CEHI_Dis_m := DisFromHIAvg_m;
DisDiff_m := DisFromH_m - DisFromI_m;

DeltaCH_CE_deg := F_Norm180(Ang_deg := (ThetaCH_rad - thetaCE_rad) * RAD2DEG_local);

// 检查量
CE_L_Check_m := SQRT((Ex - Cx) * (Ex - Cx) + (Ez - Cz) * (Ez - Cz));

Q_Offset_Check_m := SQRT(
    (Dx - Qx) * (Dx - Qx) +
    (Dz - Qz) * (Dz - Qz)
);

CH_L_Check_m := SQRT(
    (Hx - Cx) * (Hx - Cx) +
    (Hz - Cz) * (Hz - Cz)
);

EI_L_Check_m := SQRT(
    (Ix - Ex) * (Ix - Ex) +
    (Iz - Ez) * (Iz - Ez)
);

HI_L_Check_m := SQRT(
    (Ix - Hx) * (Ix - Hx) +
    (Iz - Hz) * (Iz - Hz)
);

HI_ParallelErr_m := SQRT(
    ((Ix - Hx) - (Ex - Cx)) * ((Ix - Hx) - (Ex - Cx)) +
    ((Iz - Hz) - (Ez - Cz)) * ((Iz - Hz) - (Ez - Cz))
);

Valid := TRUE;
ErrorID := 0;

END_FUNCTION_BLOCK

// ---- POUs/F_Atan2_LREAL.TcPOU
FUNCTION F_Atan2_LREAL : LREAL
VAR_INPUT
    y : LREAL;
    x : LREAL;
END_VAR
VAR
    PI_local : LREAL := 3.141592653589793;
END_VAR

IF x > 0.0 THEN
    F_Atan2_LREAL := ATAN(y / x);
ELSIF x < 0.0 THEN
    IF y >= 0.0 THEN
        F_Atan2_LREAL := ATAN(y / x) + PI_local;
    ELSE
        F_Atan2_LREAL := ATAN(y / x) - PI_local;
    END_IF;
ELSE
    IF y > 0.0 THEN
        F_Atan2_LREAL := PI_local / 2.0;
    ELSIF y < 0.0 THEN
        F_Atan2_LREAL := -PI_local / 2.0;
    ELSE
        F_Atan2_LREAL := 0.0;
    END_IF;
END_IF;

END_FUNCTION

// ---- POUs/F_Norm180.TcPOU
// =============================================================
// FUNCTION：F_Norm180
// =============================================================
FUNCTION F_Norm180 : LREAL
VAR_INPUT
    Ang_deg : LREAL;
END_VAR
VAR
    a : LREAL;
END_VAR



a := Ang_deg;

WHILE a > 180.0 DO
    a := a - 360.0;
END_WHILE;

WHILE a < -180.0 DO
    a := a + 360.0;
END_WHILE;

F_Norm180 := a;

END_FUNCTION

// ---- POUs/F_Calc_CAF_Angle_deg.TcPOU
// =============================================================
// FUNCTION：F_Calc_CAF_Angle_deg
// =============================================================
FUNCTION F_Calc_CAF_Angle_deg : LREAL
VAR_INPUT
    AC_Enc_deg             : LREAL;
    AF_Enc_deg             : LREAL;

    AC_EncRef_deg          : LREAL;
    AC_ThetaRef_deg        : LREAL;

    AF_HorizontalEnc_deg   : LREAL;
    GCH_Angle_deg          : LREAL;
    AF_EndOffset_deg       : LREAL;
END_VAR
VAR
    ThetaAC_deg       : LREAL;
    AF_ToolPitch_deg  : LREAL;
    AF_True_deg       : LREAL;
    diff_deg          : LREAL;
END_VAR



// AC 编码器 -> AC 真实机构角
ThetaAC_deg := AC_ThetaRef_deg - (AC_Enc_deg - AC_EncRef_deg);

// AF 编码器 -> 末端相对水平角。AF=205 水平时为 0。
AF_ToolPitch_deg := AF_HorizontalEnc_deg - AF_Enc_deg;

// AF 真实角度 = ToolPitch + ∠GCH + 末端偏置
AF_True_deg := AF_ToolPitch_deg + GCH_Angle_deg + AF_EndOffset_deg;

// ∠CAF
diff_deg := F_Norm180(Ang_deg := AF_True_deg - ThetaAC_deg);

F_Calc_CAF_Angle_deg := ABS(diff_deg);

END_FUNCTION

// ---- POUs/F_Calc_CEHI_Dis_m.TcPOU
// =============================================================
// FUNCTION：F_Calc_CEHI_Dis_m
// 与 FB_Calc_CEHI_Geo 同一模型，但只返回 H/I 到 CE 的平均距离。
// 返回 -1.0 表示几何无效。
// =============================================================
FUNCTION F_Calc_CEHI_Dis_m : LREAL
VAR_INPUT
    BD_Enc_mm             : LREAL;
    AC_Enc_deg            : LREAL;
    AF_Enc_deg            : LREAL;

    BD_KinOffset_mm       : LREAL;

    AC_EncRef_deg         : LREAL;
    AC_ThetaRef_deg       : LREAL;

    Ax0                   : LREAL;
    Az0                   : LREAL;
    Bx0                   : LREAL;
    Bz0                   : LREAL;

    l_AC_m                : LREAL;
    l_CD_m                : LREAL;
    l_CE_m                : LREAL;
    qOffset_m             : LREAL;
    l_CH_m                : LREAL;

    BD_BRANCH             : LREAL;
    CE_SIGN               : LREAL;

    AF_HorizontalEnc_deg  : LREAL;
    AF_CHOffset_deg       : LREAL;
    AF_EncDir_CH          : LREAL;

    GeoMargin_m           : LREAL;
END_VAR
VAR
    LBD_m        : LREAL;

    ThetaAC_deg  : LREAL;
    ThetaAC_rad  : LREAL;

    Cx_f         : LREAL;
    Cz_f         : LREAL;
    Dx_f         : LREAL;
    Dz_f         : LREAL;
    Ex_f         : LREAL;
    Ez_f         : LREAL;
    Hx_f         : LREAL;
    Hz_f         : LREAL;
    Ix_f         : LREAL;
    Iz_f         : LREAL;

    dxBC_f       : LREAL;
    dzBC_f       : LREAL;
    dBC_f        : LREAL;

    alphaBC_f    : LREAL;
    cosBeta_f    : LREAL;
    beta_f       : LREAL;
    thBD_f       : LREAL;

    thetaCD_f    : LREAL;
    thetaCE_f    : LREAL;

    s_CD_CE_f    : LREAL;
    gamma_DCE_f  : LREAL;

    uCEx_f       : LREAL;
    uCEz_f       : LREAL;
    uCHx_f       : LREAL;
    uCHz_f       : LREAL;

    thetaCH_deg  : LREAL;
    thetaAF_abs_deg : LREAL;
    thetaCH_rad  : LREAL;

    DisH_f       : LREAL;
    DisI_f       : LREAL;

    GCH_Matlab_deg : LREAL := 90.0;
    DEG2RAD_local  : LREAL := 0.0174532925199433;
END_VAR


// 默认 -1 表示几何无效
F_Calc_CEHI_Dis_m := -1.0;

// BD 编码器 -> 实际机构长度
LBD_m := (BD_Enc_mm + BD_KinOffset_mm) / 1000.0;

// AC 编码器 -> AC 机构角
ThetaAC_deg := AC_ThetaRef_deg - (AC_Enc_deg - AC_EncRef_deg);
ThetaAC_rad := ThetaAC_deg * DEG2RAD_local;

// C 点
Cx_f := Ax0 + l_AC_m * COS(ThetaAC_rad);
Cz_f := Az0 + l_AC_m * SIN(ThetaAC_rad);

// B-C
dxBC_f := Cx_f - Bx0;
dzBC_f := Cz_f - Bz0;
dBC_f  := SQRT(dxBC_f * dxBC_f + dzBC_f * dzBC_f);

IF (LBD_m <= 0.01) OR (dBC_f <= 0.01) THEN
    RETURN;
END_IF;
//三角形存在性判断
IF NOT ((dBC_f < (LBD_m + l_CD_m - GeoMargin_m)) AND
        (dBC_f > (ABS(LBD_m - l_CD_m) + GeoMargin_m))) THEN
    RETURN;//理论边界预留安全余量
END_IF;

// 三角形 B-C-D求解
alphaBC_f := F_Atan2_LREAL(y := dzBC_f, x := dxBC_f);

cosBeta_f := (LBD_m * LBD_m + dBC_f * dBC_f - l_CD_m * l_CD_m)
             / (2.0 * LBD_m * dBC_f);

IF cosBeta_f > 1.0 THEN
    cosBeta_f := 1.0;
ELSIF cosBeta_f < -1.0 THEN
    cosBeta_f := -1.0;
END_IF;//数值鲁棒处理防止accos越界

beta_f := ACOS(cosBeta_f);
thBD_f := alphaBC_f + BD_BRANCH * beta_f;

Dx_f := Bx0 + LBD_m * COS(thBD_f);
Dz_f := Bz0 + LBD_m * SIN(thBD_f);

thetaCD_f := F_Atan2_LREAL(y := Dz_f - Cz_f, x := Dx_f - Cx_f);

// D 到 CE 的垂直偏置 qOffset_m
IF l_CD_m <= ABS(qOffset_m) THEN
    RETURN;
END_IF;

s_CD_CE_f   := SQRT(l_CD_m * l_CD_m - qOffset_m * qOffset_m);
gamma_DCE_f := ATAN(qOffset_m / s_CD_CE_f);

thetaCE_f := thetaCD_f + CE_SIGN * gamma_DCE_f;

uCEx_f := COS(thetaCE_f);
uCEz_f := SIN(thetaCE_f);

Ex_f := Cx_f + l_CE_m * uCEx_f;
Ez_f := Cz_f + l_CE_m * uCEz_f;

// MATLAB 后级 H/I 方法,一致性，无实际意义
thetaCH_deg := AF_EncDir_CH * (AF_Enc_deg - AF_HorizontalEnc_deg) + AF_CHOffset_deg;
thetaAF_abs_deg := thetaCH_deg + GCH_Matlab_deg;
thetaCH_deg := thetaAF_abs_deg - GCH_Matlab_deg;
thetaCH_rad := thetaCH_deg * DEG2RAD_local;

uCHx_f := COS(thetaCH_rad);
uCHz_f := SIN(thetaCH_rad);

Hx_f := Cx_f + l_CH_m * uCHx_f;
Hz_f := Cz_f + l_CH_m * uCHz_f;

Ix_f := Ex_f + (Hx_f - Cx_f);
Iz_f := Ez_f + (Hz_f - Cz_f);

DisH_f := ABS(
    uCEx_f * (Hz_f - Cz_f) - uCEz_f * (Hx_f - Cx_f)
);

DisI_f := ABS(
    uCEx_f * (Iz_f - Cz_f) - uCEz_f * (Ix_f - Cx_f)
);

F_Calc_CEHI_Dis_m := 0.5 * (DisH_f + DisI_f);

END_FUNCTION

// ---- POUs/F_CEHI_CandidateAllow.TcPOU
// =============================================================
// FUNCTION：F_CEHI_CandidateAllow
// 逐方向预测放行逻辑。
// =============================================================
FUNCTION F_CEHI_CandidateAllow : BOOL
VAR_INPUT
    CurrentValid   : BOOL;
    CurrentDis_m   : LREAL;
    CandidateDis_m : LREAL;
    MinSafe_m      : LREAL;
    ImproveEps_m   : LREAL;
END_VAR



F_CEHI_CandidateAllow := FALSE;

IF CandidateDis_m <= 0.0 THEN
    RETURN;
END_IF;

IF CurrentValid THEN
    IF CurrentDis_m < MinSafe_m THEN
        // 已经小于安全边界：只允许让距离增大的方向。
        F_CEHI_CandidateAllow := CandidateDis_m > (CurrentDis_m + ImproveEps_m);
    ELSE
        // 尚未越界：允许在安全边界以上运动，包括距离变小但不越界。
        F_CEHI_CandidateAllow := CandidateDis_m >= MinSafe_m;
    END_IF;
ELSE
    // 当前几何无效：只允许候选回到安全边界以上。
    F_CEHI_CandidateAllow := CandidateDis_m >= MinSafe_m;
END_IF;

END_FUNCTION

// ---- POUs/F_Atan2_LR.TcPOU
FUNCTION F_Atan2_LR : LREAL
VAR_INPUT
    y : LREAL;
    x : LREAL;
END_VAR
VAR
    PI : LREAL := 3.14159265358979323846;
END_VAR


IF x > 1.0E-12 THEN
    F_Atan2_LR := ATAN(y / x);
ELSIF x < -1.0E-12 THEN
    IF y >= 0.0 THEN
        F_Atan2_LR := ATAN(y / x) + PI;
    ELSE
        F_Atan2_LR := ATAN(y / x) - PI;
    END_IF;
ELSE
    IF y > 1.0E-12 THEN
        F_Atan2_LR := PI * 0.5;
    ELSIF y < -1.0E-12 THEN
        F_Atan2_LR := -PI * 0.5;
    ELSE
        F_Atan2_LR := 0.0;
    END_IF;
END_IF;

END_FUNCTION
